FUNCTION_BLOCK TcoKukaKss_StartProgramTask_v_9_3_x EXTENDS TcoKukaKssTask_v_9_3_x
VAR
	_stopType : TcoAbstractions.eTcoRoboticsStopType;
END_VAR

IF Execute() THEN
	_blink(inOnTime:=T#500MS,inOffTime:=T#500MS);

	IF _progress = 0 THEN
		IF CheckReferences() THEN
			_progress := _progress + 1;
		END_IF
	END_IF

	IF _progress = 1 THEN
		// AX step 0: waiting for 'InterfaceActivated'
		inoControl.ActivateInterface := TRUE;
		_varInfo :=__VARINFO(inoStatus.State.InterfaceActivated);
		THIS^.Messenger.OnCondition(_infoTimer.Q AND NOT inoStatus.State.InterfaceActivated).Warning(_sb.Clear().Append('<#Waiting for signal: #>').Append(_varInfo.Symbol).ToString());
		IF inoStatus.State.InterfaceActivated THEN
			_progress := _progress + 1;
		END_IF
	END_IF

	IF _progress = 2 THEN
		// as AX step 1, but waits for 'DrivesReady' instead of switching the drives on
		inoControl.MoveEnable := TRUE;
		inoControl.DrivesOff := TRUE;
		inoControl.ActionNo := 255;
		inoControl.ErrorConfirmation := inoStatus.State.StopMess AND NOT _blink.outQ;
		_varInfo :=__VARINFO(inoStatus.State.DrivesReady);
		THIS^.Messenger.OnCondition(_infoTimer.Q AND NOT inoStatus.State.DrivesReady).Warning(_sb.Clear().Append('<#Waiting for signal: #>').Append(_varInfo.Symbol).ToString());
		IF inoStatus.State.DrivesReady THEN
			_progress := _progress + 1;
		END_IF
	END_IF

	IF _progress = 3 THEN
		// AX step 4: acknowledge, waiting for 'StopMess' to be off
		inoControl.ErrorConfirmation := inoStatus.State.StopMess AND _blink.outQ;
		_varInfo :=__VARINFO(inoStatus.State.StopMess);
		THIS^.Messenger.OnCondition(_infoTimer.Q AND inoStatus.State.StopMess).Warning(_sb.Clear().Append('<#Waiting for signal: #>').Append(_varInfo.Symbol).Append('<# is OFF#>').ToString());
		IF NOT inoStatus.State.StopMess THEN
			_progress := _progress + 1;
		END_IF
	END_IF

	IF _progress = 4 THEN
		// AX step 5: waiting for 'RcReady'
		inoControl.MoveEnable := TRUE;
		inoControl.ErrorConfirmation := inoStatus.State.AlarmStopActive AND NOT _blink.outQ;
		_varInfo :=__VARINFO(inoStatus.State.RcReady);
		THIS^.Messenger.OnCondition(_infoTimer.Q AND NOT inoStatus.State.RcReady).Warning(_sb.Clear().Append('<#Waiting for signal: #>').Append(_varInfo.Symbol).ToString());
		IF inoStatus.State.RcReady THEN
			_progress := _progress + 1;
		END_IF
	END_IF

	IF _progress = 5 THEN
		// AX step 6: external start, waiting for 'ProActive'
		IF inoStatus.State.StopMess OR NOT inoStatus.State.RcReady OR inoStatus.State.NormalStop THEN
			inoControl.ExternalStart := FALSE; // not in AX: do not leave EXT_START high while the sequence restarts
			_progress := 1;
		ELSE
			inoControl.ExternalStart := _blink.outQ;
			_varInfo :=__VARINFO(inoStatus.State.ProActive);
			THIS^.Messenger.OnCondition(_infoTimer.Q AND NOT inoStatus.State.ProActive).Warning(_sb.Clear().Append('<#Waiting for program running signal! #>').Append(_varInfo.Symbol).ToString());
			IF inoStatus.State.ProActive THEN
				inoControl.ExternalStart := FALSE;
				_progress := _progress + 1;
			END_IF
		END_IF
	END_IF

	IF _progress = 6 THEN
		DoneWhen(TRUE);
	END_IF

	CallTimers(TRUE);
	THIS^.ThrowWhen(_errorTimer.Q);
END_IF

IF THIS^.Error AND NOT _errorMessage.Pinned THEN
	THIS^.Restore();
END_IF

METHOD INTERNAL InvokeWithParams : ITcoTaskStatus
VAR_INPUT
	inStopType : eTcoRoboticsStopType;
END_VAR
_stopType := inStopType;
InvokeWithParams := THIS^.Invoke();
END_METHOD

METHOD PUBLIC FB_init : BOOL
VAR_INPUT
    bInitRetains : BOOL; // if TRUE, the retain variables are initialized (warm start / cold start)
    bInCopyCode : BOOL; // if TRUE, the instance afterwards gets moved into the copy code (online change)
    ParentObject : ITcoObject;
END_VAR
END_METHOD

(*~
	<docu>
		<summary>
			Executes when task is aborted.
		</summary>			
	</docu>	
~*)
METHOD PROTECTED OnAbort
IF __ISVALIDREF(inoStatus) THEN THIS^.inoStatus.ActionDescription := '<#Start program was aborted.#>'; END_IF;
IF __ISVALIDREF(inoControl) THEN
	inoControl.ExternalStart := FALSE;
	inoControl.ErrorConfirmation := FALSE;
	inoControl.MoveEnable := FALSE;
END_IF
END_METHOD

(*~
	<docu>
		<summary>
			Executes when task reaches the ```Done``` state .
		</summary>			
	</docu>	
~*)
METHOD PROTECTED OnDone
IF __ISVALIDREF(inoStatus) THEN THIS^.inoStatus.ActionDescription := '<#Start program finished successfully.#>'; END_IF;
_progress := 0;
END_METHOD

(*~
	<docu>
		<summary>
			Executes when task reaches the ```Error``` state.
		</summary>			
	</docu>	
~*)
METHOD PROTECTED OnError
VAR
	description: STRING;
END_VAR
description := '<#Start program finished with error.#>';
IF __ISVALIDREF(inoStatus) THEN THIS^.inoStatus.ActionDescription := description; END_IF;
THIS^._errorMessage.Error(_sb.Clear().Append(description).Append(' To restore acknowledge this alarm.').ToString()).Pin();
IF __ISVALIDREF(inoControl) THEN
	inoControl.ExternalStart := FALSE;
END_IF
END_METHOD

METHOD PROTECTED OnStart
IF __ISVALIDREF(inoStatus) THEN THIS^.inoStatus.ActionDescription := '<#Start program started.#>'; END_IF;
CallTimers(FALSE);
IF __ISVALIDREF(inoControl) THEN
	inoControl.ExternalStart := FALSE;
	inoControl.ActivateInterface := FALSE;
END_IF
END_METHOD

(*~
	<docu>
		<summary>
			Restores this instance to the Ready state. Can be called explicitly or from within one of the restore mechanisms.
			<para>
				See also <see cref="PlcDocu.TcoCore.TcoTask.AutoRestorable()"/>
			</para>
		</summary>
	</docu>
~*)
METHOD Restore : ITcoRestorable
SUPER^.Restore();
END_METHOD

END_FUNCTION_BLOCK

(* stored: Version 1.1.0.1, ProductVersion 3.1.4024.12
   POU TcoKukaKss_StartProgramTask_v_9_3_x: Id {e88a169f-bd92-488f-a4da-aa4fb8870a16}, SpecialFunc None
   Method InvokeWithParams: Id {90e1d21f-2fdd-45e2-b8bb-47356c40529d}
   Method FB_init: Id {54ca6f24-512b-46d3-9368-a507c8d7f253}
   Method OnAbort: Id {e2e482d0-adbd-4112-9a36-399ed0b2a8b0}
   Method OnDone: Id {3325cf26-3d6a-40a2-a054-7d85736b5780}
   Method OnError: Id {c9cc5a16-982f-463d-8e69-11e0cca96b3d}
   Method OnStart: Id {17c51b7f-2d05-4a25-b964-6d4188921f88}
   Method Restore: Id {29f429be-cc7d-4639-8077-301a2e1b2622} *)
